SUBAPPLICATION Uebung_159b (* Übung zu FsServer: Datei zum logiBUS-File-Server schicken (Gerät A) *)
  (* Standard: 61499-2; Description: Copyright (c) 2026 Meisterschulen am Ostbahnhof This program and the accompanying materials are made available under the terms of the Eclipse Public License 2.0 which is available at https://www.eclipse.org/legal/epl-2.0/ SPDX-License-Identifier: EPL-2.0 *)
  (* Version 1.0, 2026-11-26, Franz Höpfinger, Meisterschulen am Ostbahnhof, initial API and implementation and/or initial documentation *)
  PACKAGE Uebungen;
  IMPORT Uebungen::const::Uebung_150_159::FileServer::FS_ADD_LOGIBUS;
  IMPORT Uebungen::const::Uebung_150_159::FileServer::FS_FLT_LOGIBUS;
  IMPORT Uebungen::const::Uebung_150_159::FileServer::FS_LOGIBUS_DATEI;
  IMPORT Uebungen::const::Uebung_150_159::FileServer::FS_LOGIBUS_ORDNER;
  IMPORT Uebungen::const::Uebung_150_159::FileServer::FS_LOKAL;
  IMPORT Uebungen::const::Uebung_150_159::FileServer::FS_LOKAL_ZURUECK;
  IMPORT isobus::pgn::ISOUSERHOME_e::network;
  IMPORT isobus::pgn::ISO_CAN_NODE::NODE1;
  IMPORT logiBUS::io::DI::logiBUS_DI::Input_I1;
  IMPORT logiBUS::io::DI::logiBUS_DI_Events::BUTTON_SINGLE_CLICK;
  IMPORT logiBUS::io::DQ::logiBUS_DO::Output_Q1;
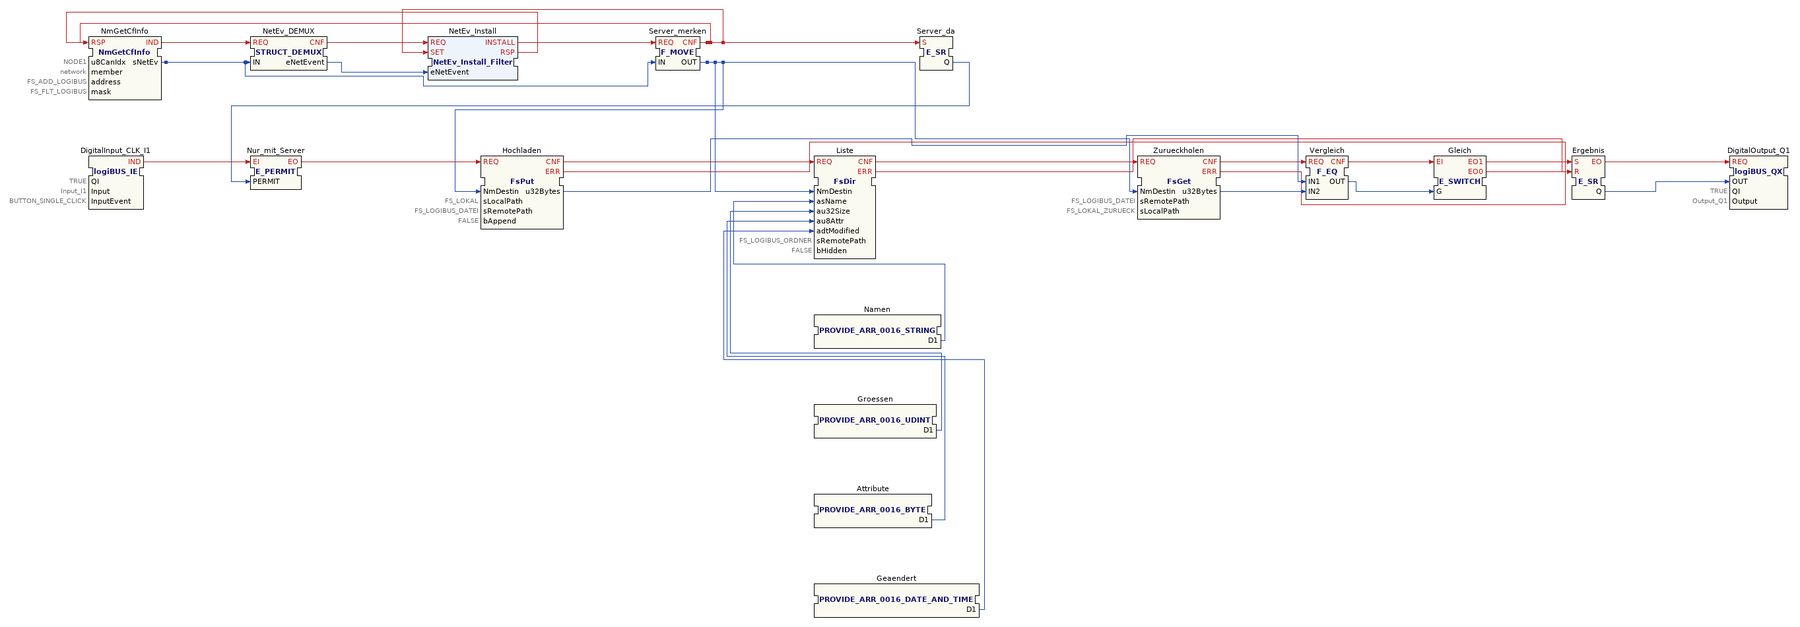
  (* Datei zum logiBUS-File-Server schicken (FsPut, FsDir, FsGet), Gerät A. Gegenstück: Übung 159 auf Gerät B. NmGetCfInfo filtert auf NAME-Funktion 61 UND Herstellercode 1116 (FS_ADD_LOGIBUS/FS_FLT_LOGIBUS), sonst käme der File Server des Terminals. I1 Klick (nur mit Server): FS_LOKAL nach \\LOGIBUS\IMPORT\test.txt, Ordner listen, Datei nach FS_LOKAL_ZURUECK zurückholen, Bytes vergleichen. Q1 an = gleich. Pfade am Server immer mit Volume: B hat ohne Stick kein Primary Volume, relative Pfade gehen ins Leere. FS_LOKAL muss es geben (Übung 156b). Watch: Liste.asName/u16Count, Hochladen.u32Bytes, Zurueckholen.u32Bytes; bei ERR s16Status und u16FsError (8 = Quota voll). Voraussetzungen: PART_13_FSC = 1 in /data/functionalities.ini, Firmware mit File Server, neue isobus_fs-ELF. *)
  FBS
    NmGetCfInfo : isobus::pgn::NmGetCfInfo(u8CanIdx := NODE1, member := network, address := FS_ADD_LOGIBUS, mask := FS_FLT_LOGIBUS); (* meldet nur den logiBUS-File-Server (Funktion 61, Hersteller 1116) *)
    NetEv_DEMUX : eclipse4diac::convert::STRUCT_DEMUX; {SET_ATTRIBUTE(StructuredType, isobus::pgn::ISONETEVENT_T)}
    Server_merken : iec61131::selection::F_MOVE; (* eigener CF und File-Server-CF (NmDestin) *)
    Server_da : iec61499::events::E_SR;
    DigitalInput_CLK_I1 : logiBUS::io::DI::logiBUS_IE(QI := TRUE, Input := Input_I1, InputEvent := BUTTON_SINGLE_CLICK);
    Nur_mit_Server : iec61499::events::E_PERMIT;
    Hochladen : isobus::fs::FsPut(sLocalPath := FS_LOKAL, sRemotePath := FS_LOGIBUS_DATEI, bAppend := FALSE); (* FS_LOKAL nach \\LOGIBUS\IMPORT\test.txt (mit Volume!) *)
    Namen : eclipse4diac::convert::providers::PROVIDE_ARR_0016_STRING;
    Groessen : eclipse4diac::convert::providers::PROVIDE_ARR_0016_UDINT;
    Attribute : eclipse4diac::convert::providers::PROVIDE_ARR_0016_BYTE;
    Geaendert : eclipse4diac::convert::providers::PROVIDE_ARR_0016_DATE_AND_TIME;
    Liste : isobus::fs::FsDir(sRemotePath := FS_LOGIBUS_ORDNER, bHidden := FALSE); (* \\LOGIBUS\IMPORT listen (test.txt muss dabei sein) *)
    Zurueckholen : isobus::fs::FsGet(sRemotePath := FS_LOGIBUS_DATEI, sLocalPath := FS_LOKAL_ZURUECK); (* test.txt nach FS_LOKAL_ZURUECK holen *)
    Vergleich : iec61131::comparison::F_EQ; (* gleich viele Bytes hin und zurück? *)
    Gleich : iec61499::events::E_SWITCH;
    Ergebnis : iec61499::events::E_SR; (* Q1 an = hin und zurück gleich groß *)
    DigitalOutput_Q1 : logiBUS::io::DQ::logiBUS_QX(QI := TRUE, Output := Output_Q1);
  END_FBS
  SUBAPPS
    NetEv_Install : MyLib::sys::NetEv_Install_Filter;
  END_SUBAPPS
  EVENT_CONNECTIONS
    NmGetCfInfo.IND TO NetEv_DEMUX.REQ;
    NetEv_DEMUX.CNF TO NetEv_Install.REQ;
    NetEv_Install.INSTALL TO Server_merken.REQ;
    NetEv_Install.RSP TO NmGetCfInfo.RSP;
    Server_merken.CNF TO NetEv_Install.SET;
    Server_merken.CNF TO Server_da.S;
    Server_merken.CNF TO NmGetCfInfo.RSP;
    DigitalInput_CLK_I1.IND TO Nur_mit_Server.EI;
    Nur_mit_Server.EO TO Hochladen.REQ;
    Hochladen.CNF TO Liste.REQ;
    Liste.CNF TO Zurueckholen.REQ;
    Zurueckholen.CNF TO Vergleich.REQ;
    Vergleich.CNF TO Gleich.EI;
    Gleich.EO1 TO Ergebnis.S;
    Gleich.EO0 TO Ergebnis.R;
    Hochladen.ERR TO Ergebnis.R;
    Liste.ERR TO Ergebnis.R;
    Zurueckholen.ERR TO Ergebnis.R;
    Ergebnis.EO TO DigitalOutput_Q1.REQ;
  END_CONNECTIONS
  DATA_CONNECTIONS
    NmGetCfInfo.sNetEv TO NetEv_DEMUX.IN;
    NetEv_DEMUX.eNetEvent TO NetEv_Install.eNetEvent;
    NmGetCfInfo.sNetEv TO Server_merken.IN;
    Server_merken.OUT TO Hochladen.NmDestin;
    Server_merken.OUT TO Liste.NmDestin;
    Server_merken.OUT TO Zurueckholen.NmDestin;
    Namen.D1 TO Liste.asName;
    Groessen.D1 TO Liste.au32Size;
    Attribute.D1 TO Liste.au8Attr;
    Geaendert.D1 TO Liste.adtModified;
    Hochladen.u32Bytes TO Vergleich.IN1;
    Zurueckholen.u32Bytes TO Vergleich.IN2;
    Vergleich.OUT TO Gleich.G;
    Server_da.Q TO Nur_mit_Server.PERMIT;
    Ergebnis.Q TO DigitalOutput_Q1.OUT;
  END_CONNECTIONS
END_SUBAPPLICATION
